(* IEC 61131-3 sources: ConveyorControl-with-PLC/4E_Gruppe1_Graf_Projekt1/Network, 1 file *)

(* ---- ConfigObjects.st ---- *)
FUNCTION GLOBAL TAB TASK_CONF
_K_TASK, _K_REAL,
_K_END_VAR,

_K_TASK, _K_CYCLIC,
_K_END_VAR,

_K_TASK, _K_BACKGROUND,
_K_END_VAR,

_K_END_CONF
END_FUNCTION

FUNCTION GLOBAL TAB IPR_CONF
_K_IPR
	0$UINT,
_K_END_VAR,
_K_END_CONF
END_FUNCTION

FUNCTION GLOBAL TAB CONFIG_TABLES
00058$UINT,
0$UINT, 1, 7, "_BUSINTERFACESDIASDRIVEMNG",
0$UINT, 1, 58, "_DRIVEAXIS",
0$UINT, 1, 67, "_DRIVEAXISBASE",
0$UINT, 1, 20, "_DRIVEAXISSET",
0$UINT, 1, 7, "_DRIVEMNG_DC062",
0$UINT, 1, 54, "_DRIVEMNG_MDD100",
0$UINT, 1, 39, "_DRIVEMNGBASE",
0$UINT, 1, 18, "_FILESYS",
0$UINT, 0, 1, "_LINKER",
0$UINT, 1, 1, "_MULTITASK",
0$UINT, 0, 4, "_OSKERNEL",
0$UINT, 0, 0, "_STDLIB",
0$UINT, 1, 1, "_TASKOBJECTCONTROL",
0$UINT, 1, 58, "_VARANDRIVEBASE",
0$UINT, 0, 0, "ABSCHLUSS",
0$UINT, 1, 27, "AM441",
0$UINT, 1, 17, "BUSINTERFACESDIAS",
0$UINT, 1, 27, "BUSINTERFACESDIASINTERNAL",
0$UINT, 0, 0, "CLASS0",
0$UINT, 1, 36, "DI200",
0$UINT, 2, 32, "DIASMASTER",
0$UINT, 1, 75, "DIASMASTERC",
0$UINT, 2, 15, "DIASMASTERMAIN",
0$UINT, 1, 0, "DIASMASTERPOSTSCAN",
0$UINT, 1, 11, "EEPROM",
0$UINT, 1, 20, "HUB_BASE",
0$UINT, 2, 10, "HUB_BASE_ROOT",
0$UINT, 2, 31, "HWBASE",
0$UINT, 2, 51, "HWBASECDIAS",
0$UINT, 4, 0, "HWCONTROL",
0$UINT, 1, 10, "HWCONTROLBASE",
0$UINT, 1, 0, "HWRTPOSTSCAN",
0$UINT, 1, 6, "I2CCDIAS",
0$UINT, 1, 21, "MERKEREX",
0$UINT, 1, 16, "RAMEX",
0$UINT, 1, 9, "RAMFILE",
0$UINT, 1, 22, "SAFETYBASE",
0$UINT, 3, 3, "SAFETYCDIAS_BASE",
0$UINT, 2, 0, "SAFETYMANAGER",
0$UINT, 1, 31, "SCP011",
0$UINT, 1, 51, "SDIASBASE",
0$UINT, 1, 10, "SDIASHUBBASE",
0$UINT, 1, 75, "SDIASMANAGER",
0$UINT, 1, 38, "SDIASPLC",
0$UINT, 1, 6, "SDIASSAFETYBASE",
0$UINT, 1, 25, "SDIASSAFETYMANAGER",
0$UINT, 1, 4, "SDM081",
0$UINT, 1, 10, "STRING",
0$UINT, 1, 80, "STRINGINTERNAL",
0$UINT, 1, 20, "SYNCCALL",
0$UINT, 1, 38, "TO127",
0$UINT, 2, 7, "VARAN_BASE",
0$UINT, 2, 26, "VARANMANAGER",
0$UINT, 1, 68, "VARANMANAGER_2",
0$UINT, 1, 21, "VARANMANAGER_BASE",
0$UINT, 1, 1, "VARANMANAGERPOSTSCAN",
0$UINT, 1, 3, "VIRTUALBASEINIT",
0$UINT, 2, 10, "WATCHDOGDIAS",
ONE_CFG$UINT, 0, 0, "ONE_HW_Network",
ONE_CFG$UINT, 0, 0, "ONE_net0",
TASK_CFG$UINT, 0, 0, "TASK_CONF",
IPR_CFG$UINT, 0, 0, "IPR_CONF",
PRJ_CFG$UINT, 0, 0, "4E_Gruppe1_Graf_Projekt1",
END_FUNCTION

#ifdef __LSLLDR_IOELEMENTS__
FUNCTION GLOBAL TAB _IO_ELEMENTS_TAB
0000$UINT, 0005$UINT,
"**IOCONN_EMPTY**", "_DriveAxis1.AxEnable",
"IO_Element0", "DI2001.Input1",
"IO_Element1", "DI2001.Input2",
"IO_Element2", "TO1271.Output1",
"IO_Element3", "TO1271.Output2",
END_FUNCTION
#endif //__LSLLDR_IOELEMENTS__
